(* IEC 61131-3 sources: smart-manufacture/PART06, 11 files *)

(* ---- ld1_sensor.st ---- *)
PROGRAM conveyor
  VAR
    RAW_A    AT %IX0.3 : BOOL;     (* 센서 A 원래 값  GPIO17 · 물리 11번 *)
    RAW_B    AT %IX0.4 : BOOL;     (* 센서 B 원래 값  GPIO27 · 물리 13번 *)
    SENSOR_A AT %QX1.3 : BOOL;     (* 센서 A  1 = 감지 (렁 0 에서 뒤집음) *)
    SENSOR_B AT %QX1.4 : BOOL;     (* 센서 B  1 = 감지 *)
    MOVE_RIGHT AT %QX0.2 : BOOL;  (* 정방향  GPIO23 · 물리 16번 = IN1 *)
    MOVE_LEFT  AT %QX0.3 : BOOL;  (* 역방향  GPIO24 · 물리 18번 = IN2 *)
  END_VAR
  (* 0 : 센서 뒤집기 — D0 는 감지 = 0 이므로 NOT 으로 1 = 감지 *)
  SENSOR_A := NOT RAW_A;
  SENSOR_B := NOT RAW_B;
  (* 1 : 센서 A 가 박스를 보는 동안만 정방향 *)
  MOVE_RIGHT := SENSOR_A;
END_PROGRAM

CONFIGURATION Config0
  RESOURCE Res0 ON PLC
    TASK task0(INTERVAL := T#50ms, PRIORITY := 0);
    PROGRAM instance0 WITH task0 : conveyor;
  END_RESOURCE
END_CONFIGURATION

(* ---- ld2_selfhold.st ---- *)
PROGRAM conveyor
  VAR
    RAW_A    AT %IX0.3 : BOOL;     (* 센서 A 원래 값  GPIO17 · 물리 11번 *)
    RAW_B    AT %IX0.4 : BOOL;     (* 센서 B 원래 값  GPIO27 · 물리 13번 *)
    SENSOR_A AT %QX1.3 : BOOL;     (* 센서 A  1 = 감지 (렁 0 에서 뒤집음) *)
    SENSOR_B AT %QX1.4 : BOOL;     (* 센서 B  1 = 감지 *)
    MOVE_RIGHT AT %QX0.2 : BOOL;  (* 정방향  GPIO23 · 물리 16번 = IN1 *)
    MOVE_LEFT  AT %QX0.3 : BOOL;  (* 역방향  GPIO24 · 물리 18번 = IN2 *)
  END_VAR
  (* 0 : 센서 뒤집기 — D0 는 감지 = 0 이므로 NOT 으로 1 = 감지 *)
  SENSOR_A := NOT RAW_A;
  SENSOR_B := NOT RAW_B;
  (* 1 : 센서 A 가 한 번 보면 계속 정방향 (자기유지) *)
  MOVE_RIGHT := SENSOR_A OR MOVE_RIGHT;
END_PROGRAM

CONFIGURATION Config0
  RESOURCE Res0 ON PLC
    TASK task0(INTERVAL := T#50ms, PRIORITY := 0);
    PROGRAM instance0 WITH task0 : conveyor;
  END_RESOURCE
END_CONFIGURATION

(* ---- ld3_break.st ---- *)
PROGRAM conveyor
  VAR
    RAW_A    AT %IX0.3 : BOOL;     (* 센서 A 원래 값  GPIO17 · 물리 11번 *)
    RAW_B    AT %IX0.4 : BOOL;     (* 센서 B 원래 값  GPIO27 · 물리 13번 *)
    SENSOR_A AT %QX1.3 : BOOL;     (* 센서 A  1 = 감지 (렁 0 에서 뒤집음) *)
    SENSOR_B AT %QX1.4 : BOOL;     (* 센서 B  1 = 감지 *)
    MOVE_RIGHT AT %QX0.2 : BOOL;  (* 정방향  GPIO23 · 물리 16번 = IN1 *)
    MOVE_LEFT  AT %QX0.3 : BOOL;  (* 역방향  GPIO24 · 물리 18번 = IN2 *)
  END_VAR
  (* 0 : 센서 뒤집기 — D0 는 감지 = 0 이므로 NOT 으로 1 = 감지 *)
  SENSOR_A := NOT RAW_A;
  SENSOR_B := NOT RAW_B;
  (* 1 : 자기유지 + 센서 B 의 b 접점으로 끊기 *)
  MOVE_RIGHT := (SENSOR_A OR MOVE_RIGHT) AND NOT SENSOR_B;
END_PROGRAM

CONFIGURATION Config0
  RESOURCE Res0 ON PLC
    TASK task0(INTERVAL := T#50ms, PRIORITY := 0);
    PROGRAM instance0 WITH task0 : conveyor;
  END_RESOURCE
END_CONFIGURATION

(* ---- ld4_cycle.st ---- *)
PROGRAM conveyor
  VAR
    RAW_A    AT %IX0.3 : BOOL;     (* 센서 A 원래 값  GPIO17 · 물리 11번 *)
    RAW_B    AT %IX0.4 : BOOL;     (* 센서 B 원래 값  GPIO27 · 물리 13번 *)
    SENSOR_A AT %QX1.3 : BOOL;     (* 센서 A  1 = 감지 (렁 0 에서 뒤집음) *)
    SENSOR_B AT %QX1.4 : BOOL;     (* 센서 B  1 = 감지 *)
    MOVE_RIGHT AT %QX0.2 : BOOL;  (* 정방향  GPIO23 · 물리 16번 = IN1 *)
    MOVE_LEFT  AT %QX0.3 : BOOL;  (* 역방향  GPIO24 · 물리 18번 = IN2 *)
  END_VAR
  (* 0 : 센서 뒤집기 — D0 는 감지 = 0 이므로 NOT 으로 1 = 감지 *)
  SENSOR_A := NOT RAW_A;
  SENSOR_B := NOT RAW_B;
  (* 1 : A 에서 출발 -> B 에 닿을 때까지 정방향 (자기유지 + 인터록) *)
  MOVE_RIGHT := (SENSOR_A OR MOVE_RIGHT) AND NOT SENSOR_B AND NOT MOVE_LEFT;
  (* 2 : B 에서 출발 -> A 에 닿을 때까지 역방향 *)
  MOVE_LEFT := (SENSOR_B OR MOVE_LEFT) AND NOT SENSOR_A AND NOT MOVE_RIGHT;
END_PROGRAM

CONFIGURATION Config0
  RESOURCE Res0 ON PLC
    TASK task0(INTERVAL := T#50ms, PRIORITY := 0);
    PROGRAM instance0 WITH task0 : conveyor;
  END_RESOURCE
END_CONFIGURATION

(* ---- ld5_delay.st ---- *)
PROGRAM conveyor
  VAR
    RAW_A    AT %IX0.3 : BOOL;     (* 센서 A 원래 값  GPIO17 · 물리 11번 *)
    RAW_B    AT %IX0.4 : BOOL;     (* 센서 B 원래 값  GPIO27 · 물리 13번 *)
    SENSOR_A AT %QX1.3 : BOOL;     (* 센서 A  1 = 감지 (렁 0 에서 뒤집음) *)
    SENSOR_B AT %QX1.4 : BOOL;     (* 센서 B  1 = 감지 *)
    MOVE_RIGHT AT %QX0.2 : BOOL;  (* 정방향  GPIO23 · 물리 16번 = IN1 *)
    MOVE_LEFT  AT %QX0.3 : BOOL;  (* 역방향  GPIO24 · 물리 18번 = IN2 *)
    A_DONE : BOOL;                 (* A 에서 3 초 기다림 끝 *)
    B_DONE : BOOL;
    TA : TON;                      (* On-Delay 타이머 *)
    TB : TON;
  END_VAR
  (* 0 : 센서 뒤집기 — D0 는 감지 = 0 이므로 NOT 으로 1 = 감지 *)
  SENSOR_A := NOT RAW_A;
  SENSOR_B := NOT RAW_B;
  (* 1 · 2 : 끝에서 3 초 재기 *)
  TA(IN := SENSOR_A, PT := T#3s);
  A_DONE := TA.Q;
  TB(IN := SENSOR_B, PT := T#3s);
  B_DONE := TB.Q;
  (* 3 · 4 : 3 초 뒤 출발 *)
  MOVE_RIGHT := (A_DONE OR MOVE_RIGHT) AND NOT SENSOR_B AND NOT MOVE_LEFT;
  MOVE_LEFT := (B_DONE OR MOVE_LEFT) AND NOT SENSOR_A AND NOT MOVE_RIGHT;
END_PROGRAM

CONFIGURATION Config0
  RESOURCE Res0 ON PLC
    TASK task0(INTERVAL := T#50ms, PRIORITY := 0);
    PROGRAM instance0 WITH task0 : conveyor;
  END_RESOURCE
END_CONFIGURATION

(* ---- ld6_count.st ---- *)
PROGRAM conveyor
  VAR
    RAW_A    AT %IX0.3 : BOOL;     (* 센서 A 원래 값  GPIO17 · 물리 11번 *)
    RAW_B    AT %IX0.4 : BOOL;     (* 센서 B 원래 값  GPIO27 · 물리 13번 *)
    SENSOR_A AT %QX1.3 : BOOL;     (* 센서 A  1 = 감지 (렁 0 에서 뒤집음) *)
    SENSOR_B AT %QX1.4 : BOOL;     (* 센서 B  1 = 감지 *)
    MOVE_RIGHT AT %QX0.2 : BOOL;  (* 정방향  GPIO23 · 물리 16번 = IN1 *)
    MOVE_LEFT  AT %QX0.3 : BOOL;  (* 역방향  GPIO24 · 물리 18번 = IN2 *)
    A_DONE : BOOL;                 (* A 에서 3 초 기다림 끝 *)
    B_DONE : BOOL;
    TA : TON;                      (* On-Delay 타이머 *)
    TB : TON;
    CNT_RST  AT %QX2.6 : BOOL;     (* 카운트 초기화 — Monitoring 의 true · false *)
    COUNT    AT %MW0   : INT;      (* 왕복 횟수 — Monitoring 에서 보임 *)
    CNT : CTU;                     (* Up Counter — 0 → 1 될 때마다 1 씩 *)
  END_VAR
  (* 0 : 센서 뒤집기 — D0 는 감지 = 0 이므로 NOT 으로 1 = 감지 *)
  SENSOR_A := NOT RAW_A;
  SENSOR_B := NOT RAW_B;
  (* 1 : A 로 돌아올 때(MOVE_LEFT 로 가다가 A 에 닿음) 1 회 *)
  CNT(CU := SENSOR_A AND MOVE_LEFT, R := CNT_RST, PV := 9999);
  COUNT := CNT.CV;
  (* 2 · 3 : 끝에서 3 초 재기 *)
  TA(IN := SENSOR_A, PT := T#3s);
  A_DONE := TA.Q;
  TB(IN := SENSOR_B, PT := T#3s);
  B_DONE := TB.Q;
  (* 4 · 5 : 3 초 뒤 출발 *)
  MOVE_RIGHT := (A_DONE OR MOVE_RIGHT) AND NOT SENSOR_B AND NOT MOVE_LEFT;
  MOVE_LEFT := (B_DONE OR MOVE_LEFT) AND NOT SENSOR_A AND NOT MOVE_RIGHT;
END_PROGRAM

CONFIGURATION Config0
  RESOURCE Res0 ON PLC
    TASK task0(INTERVAL := T#50ms, PRIORITY := 0);
    PROGRAM instance0 WITH task0 : conveyor;
  END_RESOURCE
END_CONFIGURATION

(* ---- ld7_alarm.st ---- *)
PROGRAM conveyor
  VAR
    RAW_A    AT %IX0.3 : BOOL;     (* 센서 A 원래 값  GPIO17 · 물리 11번 *)
    RAW_B    AT %IX0.4 : BOOL;     (* 센서 B 원래 값  GPIO27 · 물리 13번 *)
    SENSOR_A AT %QX1.3 : BOOL;     (* 센서 A  1 = 감지 (렁 0 에서 뒤집음) *)
    SENSOR_B AT %QX1.4 : BOOL;     (* 센서 B  1 = 감지 *)
    MOVE_RIGHT AT %QX0.2 : BOOL;  (* 정방향  GPIO23 · 물리 16번 = IN1 *)
    MOVE_LEFT  AT %QX0.3 : BOOL;  (* 역방향  GPIO24 · 물리 18번 = IN2 *)
    A_DONE : BOOL;                 (* A 에서 3 초 기다림 끝 *)
    B_DONE : BOOL;
    TA : TON;                      (* On-Delay 타이머 *)
    TB : TON;
    CNT_RST  AT %QX2.6 : BOOL;     (* 카운트 초기화 *)
    COUNT    AT %MW0   : INT;      (* 왕복 횟수 *)
    CNT : CTU;
    ALM_RST  AT %QX2.5 : BOOL;     (* 알람 리셋 — HMI 에서도 같은 주소(코일 21) *)
    ALARM    AT %QX3.1 : BOOL;     (* 알람 — 리셋 전까지 1 유지 (코일 25) *)
    BLINK    AT %QX3.2 : BOOL;     (* 알람 깜빡임 — HMI 램프용 (코일 26) *)
    T_LOST : TON;                  (* 움직이는데 센서가 박스를 못 본 시간 *)
    T_ON : TON;                    (* 깜빡이 — 켜짐 시간 *)
    T_OFF : TON;                   (* 깜빡이 — 꺼짐 시간 *)
  END_VAR
  (* 0 : 센서 뒤집기 — D0 는 감지 = 0 이므로 NOT 으로 1 = 감지 *)
  SENSOR_A := NOT RAW_A;
  SENSOR_B := NOT RAW_B;
  (* 1 : 왕복 횟수 *)
  CNT(CU := SENSOR_A AND MOVE_LEFT, R := CNT_RST, PV := 9999);
  COUNT := CNT.CV;
  (* 2 : 모터가 도는데 10 초 동안 A · B 어느 센서도 박스를 못 보면 *)
  T_LOST(IN := (MOVE_RIGHT OR MOVE_LEFT) AND NOT SENSOR_A AND NOT SENSOR_B,
         PT := T#10s);
  (* 3 : 알람 자기유지 — ALM_RST 로만 풀림 *)
  ALARM := (T_LOST.Q OR ALARM) AND NOT ALM_RST;
  (* 4 · 5 : 끝에서 3 초 — 알람 중에는 재지 않음 *)
  TA(IN := SENSOR_A AND NOT ALARM, PT := T#3s);
  A_DONE := TA.Q;
  TB(IN := SENSOR_B AND NOT ALARM, PT := T#3s);
  B_DONE := TB.Q;
  (* 6 · 7 : 출발 — 알람이면 정지 *)
  MOVE_RIGHT := (A_DONE OR MOVE_RIGHT) AND NOT SENSOR_B
                AND NOT MOVE_LEFT AND NOT ALARM;
  MOVE_LEFT := (B_DONE OR MOVE_LEFT) AND NOT SENSOR_A
               AND NOT MOVE_RIGHT AND NOT ALARM;
  (* 8 · 9 · 10 : 알람 깜빡이 (0.5 초 켜짐 · 0.5 초 꺼짐) *)
  T_ON(IN := ALARM AND NOT T_OFF.Q, PT := T#500ms);
  T_OFF(IN := T_ON.Q, PT := T#500ms);
  BLINK := ALARM AND NOT T_ON.Q;
END_PROGRAM

CONFIGURATION Config0
  RESOURCE Res0 ON PLC
    TASK task0(INTERVAL := T#50ms, PRIORITY := 0);
    PROGRAM instance0 WITH task0 : conveyor;
  END_RESOURCE
END_CONFIGURATION

(* ---- ld8_mode.st ---- *)
PROGRAM conveyor
  VAR
    RAW_A    AT %IX0.3 : BOOL;     (* 센서 A 원래 값  GPIO17 · 물리 11번 *)
    RAW_B    AT %IX0.4 : BOOL;     (* 센서 B 원래 값  GPIO27 · 물리 13번 *)
    SENSOR_A AT %QX1.3 : BOOL;     (* 센서 A  1 = 감지 (렁 0 에서 뒤집음) *)
    SENSOR_B AT %QX1.4 : BOOL;     (* 센서 B  1 = 감지 *)
    MOVE_RIGHT AT %QX0.2 : BOOL;  (* 정방향  GPIO23 · 물리 16번 = IN1 *)
    MOVE_LEFT  AT %QX0.3 : BOOL;  (* 역방향  GPIO24 · 물리 18번 = IN2 *)
    A_DONE : BOOL;                 (* A 에서 3 초 기다림 끝 *)
    B_DONE : BOOL;
    TA : TON;                      (* On-Delay 타이머 *)
    TB : TON;
    HMI_AUTO   AT %QX2.0 : BOOL;   (* HMI 버튼 — Modbus 코일 16 *)
    HMI_MANUAL AT %QX2.1 : BOOL;   (* 코일 17 *)
    HMI_FWD    AT %QX2.2 : BOOL;   (* 수동 정방향 — 코일 18 *)
    HMI_REV    AT %QX2.3 : BOOL;   (* 수동 역방향 — 코일 19 *)
    HMI_STOP   AT %QX2.4 : BOOL;   (* 수동 정지 — 코일 20 *)
    AUTO       AT %QX3.0 : BOOL;   (* 1 = AUTO, 0 = MANUAL — 코일 24 *)
    AUTO_R : BOOL;                 (* 자동 정방향 *)
    AUTO_L : BOOL;
    MAN_R : BOOL;                  (* 수동 정방향 *)
    MAN_L : BOOL;
  END_VAR
  (* 0 : 센서 뒤집기 — D0 는 감지 = 0 이므로 NOT 으로 1 = 감지 *)
  SENSOR_A := NOT RAW_A;
  SENSOR_B := NOT RAW_B;
  (* 1 : AUTO 자기유지 — MANUAL 버튼이면 풀림 *)
  AUTO := (HMI_AUTO OR AUTO) AND NOT HMI_MANUAL;
  (* 2 · 3 : 자동 — 끝에서 3 초 *)
  TA(IN := SENSOR_A AND AUTO, PT := T#3s);
  A_DONE := TA.Q;
  TB(IN := SENSOR_B AND AUTO, PT := T#3s);
  B_DONE := TB.Q;
  (* 4 · 5 : 자동 운전 *)
  AUTO_R := (A_DONE OR AUTO_R) AND NOT SENSOR_B AND NOT AUTO_L AND AUTO;
  AUTO_L := (B_DONE OR AUTO_L) AND NOT SENSOR_A AND NOT AUTO_R AND AUTO;
  (* 6 · 7 : 수동 운전 — 끝 센서에서 스스로 멈춤 *)
  MAN_R := (HMI_FWD OR MAN_R) AND NOT HMI_STOP AND NOT SENSOR_B
           AND NOT MAN_L AND NOT AUTO;
  MAN_L := (HMI_REV OR MAN_L) AND NOT HMI_STOP AND NOT SENSOR_A
           AND NOT MAN_R AND NOT AUTO;
  (* 8 · 9 : 출력 = 자동 또는 수동 *)
  MOVE_RIGHT := (AUTO_R OR MAN_R);
  MOVE_LEFT := (AUTO_L OR MAN_L);
END_PROGRAM

CONFIGURATION Config0
  RESOURCE Res0 ON PLC
    TASK task0(INTERVAL := T#50ms, PRIORITY := 0);
    PROGRAM instance0 WITH task0 : conveyor;
  END_RESOURCE
END_CONFIGURATION

(* ---- ld9_hmi.st ---- *)
PROGRAM conveyor
  VAR
    RAW_A    AT %IX0.3 : BOOL;     (* 센서 A 원래 값  GPIO17 · 물리 11번 *)
    RAW_B    AT %IX0.4 : BOOL;     (* 센서 B 원래 값  GPIO27 · 물리 13번 *)
    SENSOR_A AT %QX1.3 : BOOL;     (* 센서 A  1 = 감지 (렁 0 에서 뒤집음) *)
    SENSOR_B AT %QX1.4 : BOOL;     (* 센서 B  1 = 감지 *)
    MOVE_RIGHT AT %QX0.2 : BOOL;  (* 정방향  GPIO23 · 물리 16번 = IN1 *)
    MOVE_LEFT  AT %QX0.3 : BOOL;  (* 역방향  GPIO24 · 물리 18번 = IN2 *)
    A_DONE : BOOL;                 (* A 에서 3 초 기다림 끝 *)
    B_DONE : BOOL;
    TA : TON;                      (* On-Delay 타이머 *)
    TB : TON;
    HMI_AUTO   AT %QX2.0 : BOOL;   (* HMI 버튼 — Modbus 코일 16 *)
    HMI_MANUAL AT %QX2.1 : BOOL;   (* 코일 17 *)
    HMI_FWD    AT %QX2.2 : BOOL;   (* 수동 정방향 — 코일 18 *)
    HMI_REV    AT %QX2.3 : BOOL;   (* 수동 역방향 — 코일 19 *)
    HMI_STOP   AT %QX2.4 : BOOL;   (* 수동 정지 — 코일 20 *)
    AUTO       AT %QX3.0 : BOOL;   (* 1 = AUTO, 0 = MANUAL — 코일 24 *)
    AUTO_R : BOOL;                 (* 자동 정방향 *)
    AUTO_L : BOOL;
    MAN_R : BOOL;                  (* 수동 정방향 *)
    MAN_L : BOOL;
    ALM_RST    AT %QX2.5 : BOOL;   (* 알람 리셋 — 코일 21 *)
    ALARM      AT %QX3.1 : BOOL;   (* 알람 — 코일 25 *)
    T_LOST : TON;                  (* 박스를 못 본 시간 *)
  END_VAR
  (* 0 : 센서 뒤집기 — D0 는 감지 = 0 이므로 NOT 으로 1 = 감지 *)
  SENSOR_A := NOT RAW_A;
  SENSOR_B := NOT RAW_B;
  (* 1 : AUTO 자기유지 — MANUAL 버튼 · 알람이면 풀림 *)
  AUTO := (HMI_AUTO OR AUTO) AND NOT HMI_MANUAL AND NOT ALARM;
  (* 2 · 3 : 자동 — 끝에서 3 초 *)
  TA(IN := SENSOR_A AND AUTO, PT := T#3s);
  A_DONE := TA.Q;
  TB(IN := SENSOR_B AND AUTO, PT := T#3s);
  B_DONE := TB.Q;
  (* 4 · 5 : 자동 운전 *)
  AUTO_R := (A_DONE OR AUTO_R) AND NOT SENSOR_B AND NOT AUTO_L AND AUTO;
  AUTO_L := (B_DONE OR AUTO_L) AND NOT SENSOR_A AND NOT AUTO_R AND AUTO;
  (* 6 · 7 : 수동 운전 — 끝 센서에서 스스로 멈춤 *)
  MAN_R := (HMI_FWD OR MAN_R) AND NOT HMI_STOP AND NOT SENSOR_B
           AND NOT MAN_L AND NOT AUTO AND NOT ALARM;
  MAN_L := (HMI_REV OR MAN_L) AND NOT HMI_STOP AND NOT SENSOR_A
           AND NOT MAN_R AND NOT AUTO AND NOT ALARM;
  (* 8 · 9 : 알람 — 프로그램 7 의 렁 2 · 3 과 같음 *)
  T_LOST(IN := (MOVE_RIGHT OR MOVE_LEFT) AND NOT SENSOR_A AND NOT SENSOR_B,
         PT := T#10s);
  ALARM := (T_LOST.Q OR ALARM) AND NOT ALM_RST;
  (* 10 · 11 : 출력 = 자동 또는 수동 *)
  MOVE_RIGHT := (AUTO_R OR MAN_R) AND NOT ALARM;
  MOVE_LEFT := (AUTO_L OR MAN_L) AND NOT ALARM;
END_PROGRAM

CONFIGURATION Config0
  RESOURCE Res0 ON PLC
    TASK task0(INTERVAL := T#50ms, PRIORITY := 0);
    PROGRAM instance0 WITH task0 : conveyor;
  END_RESOURCE
END_CONFIGURATION

(* ---- st1_cycle.st ---- *)
PROGRAM conveyor
  VAR
    RAW_A    AT %IX0.3 : BOOL;     (* 센서 A 원래 값  GPIO17 · 물리 11번 *)
    RAW_B    AT %IX0.4 : BOOL;     (* 센서 B 원래 값  GPIO27 · 물리 13번 *)
    SENSOR_A AT %QX1.3 : BOOL;     (* 센서 A  1 = 감지 (렁 0 에서 뒤집음) *)
    SENSOR_B AT %QX1.4 : BOOL;     (* 센서 B  1 = 감지 *)
    MOVE_RIGHT AT %QX0.2 : BOOL;  (* 정방향  GPIO23 · 물리 16번 = IN1 *)
    MOVE_LEFT  AT %QX0.3 : BOOL;  (* 역방향  GPIO24 · 물리 18번 = IN2 *)
  END_VAR
  (* 0 : 센서 뒤집기 — D0 는 감지 = 0 이므로 NOT 으로 1 = 감지 *)
  SENSOR_A := NOT RAW_A;
  SENSOR_B := NOT RAW_B;
  IF SENSOR_A THEN              (* A 에 닿으면 *)
    MOVE_RIGHT := TRUE;
    MOVE_LEFT := FALSE;
  ELSIF SENSOR_B THEN           (* B 에 닿으면 *)
    MOVE_RIGHT := FALSE;
    MOVE_LEFT := TRUE;
  END_IF;                       (* 둘 다 아니면 그대로 *)
END_PROGRAM

CONFIGURATION Config0
  RESOURCE Res0 ON PLC
    TASK task0(INTERVAL := T#50ms, PRIORITY := 0);
    PROGRAM instance0 WITH task0 : conveyor;
  END_RESOURCE
END_CONFIGURATION

(* ---- st2_delay.st ---- *)
PROGRAM conveyor
  VAR
    RAW_A    AT %IX0.3 : BOOL;     (* 센서 A 원래 값  GPIO17 · 물리 11번 *)
    RAW_B    AT %IX0.4 : BOOL;     (* 센서 B 원래 값  GPIO27 · 물리 13번 *)
    SENSOR_A AT %QX1.3 : BOOL;     (* 센서 A  1 = 감지 (렁 0 에서 뒤집음) *)
    SENSOR_B AT %QX1.4 : BOOL;     (* 센서 B  1 = 감지 *)
    MOVE_RIGHT AT %QX0.2 : BOOL;  (* 정방향  GPIO23 · 물리 16번 = IN1 *)
    MOVE_LEFT  AT %QX0.3 : BOOL;  (* 역방향  GPIO24 · 물리 18번 = IN2 *)
    TA : TON;
    TB : TON;
  END_VAR
  (* 0 : 센서 뒤집기 — D0 는 감지 = 0 이므로 NOT 으로 1 = 감지 *)
  SENSOR_A := NOT RAW_A;
  SENSOR_B := NOT RAW_B;
  TA(IN := SENSOR_A, PT := T#3s);
  TB(IN := SENSOR_B, PT := T#3s);
  IF TA.Q THEN                  (* A 에서 3 초 지남 -> 정방향 *)
    MOVE_RIGHT := TRUE;
    MOVE_LEFT := FALSE;
  ELSIF TB.Q THEN               (* B 에서 3 초 지남 -> 역방향 *)
    MOVE_RIGHT := FALSE;
    MOVE_LEFT := TRUE;
  ELSIF SENSOR_A OR SENSOR_B THEN   (* 끝에 막 닿음 -> 멈춤 *)
    MOVE_RIGHT := FALSE;
    MOVE_LEFT := FALSE;
  END_IF;
END_PROGRAM

CONFIGURATION Config0
  RESOURCE Res0 ON PLC
    TASK task0(INTERVAL := T#50ms, PRIORITY := 0);
    PROGRAM instance0 WITH task0 : conveyor;
  END_RESOURCE
END_CONFIGURATION
